(* IEC 61131-3 sources: Lasal-MCP/examples/SampleSource/2_PumpControlSolution/Stations/MachineControl/MachineControl/Class/PumpControl, 1 file *)

(* ---- PumpControl.st ---- *)
(*!
<Class
	Name               = "PumpControl"
	Revision           = "0.0"
	RealtimeTask       = "false"
	CyclicTask         = "true"
	DefCyclictime      = "10 ms"
	BackgroundTask     = "false"
	Sigmatek           = "false"
	OSInterface        = "false"
	HighPriority       = "false"
	Automatic          = "false"
	UpdateMode         = "Prescan"
	SharedCommandTable = "true"
	Objectsize         = "(510,360)">
	<Channels>
		<Server Name="ActFillLevelVisu" Visualized="true" Initialize="false" WriteProtected="true" Retentive="false"/>
		<Server Name="ClassSvr" Visualized="false" Initialize="false" WriteProtected="true" Retentive="false"/>
		<Server Name="MaxBorder" Visualized="true" Initialize="false" WriteProtected="false" Retentive="File"/>
		<Server Name="MinBorder" Visualized="true" Initialize="false" WriteProtected="false" Retentive="File"/>
		<Server Name="PumpVisu" Visualized="true" Initialize="false" WriteProtected="true" Retentive="false"/>
		<Client Name="ActFillLevel" Required="true" Internal="false"/>
		<Client Name="Pump" Required="true" Internal="false"/>
	</Channels>
</Class>
*)
PumpControl : CLASS
  //Servers:
	ClassSvr 	: SvrChCmd_DINT;
	MaxBorder 	: SvrCh_DINT;
	MinBorder 	: SvrCh_DINT;
	PumpVisu 	: SvrCh_DINT;
	ActFillLevelVisu 	: SvrCh_DINT;
  //Clients:
	Pump 	: CltCh_DINT;
	ActFillLevel 	: CltCh_DINT;
  //Variables:
  //Functions:

	FUNCTION VIRTUAL GLOBAL CyWork
		VAR_INPUT
			EAX 	: UDINT;
		END_VAR
		VAR_OUTPUT
			state (EAX) 	: UDINT;
		END_VAR;

	FUNCTION VIRTUAL GLOBAL PumpVisu::Read
		VAR_OUTPUT
			output (EAX) 	: DINT;
		END_VAR;

	FUNCTION VIRTUAL GLOBAL ActFillLevelVisu::Read
		VAR_OUTPUT
			output (EAX) 	: DINT;
		END_VAR;
  //Tables:
	FUNCTION @STD
		VAR_OUTPUT
			ret_code	: CONFSTATES;
		END_VAR;
	FUNCTION GLOBAL TAB @CT_;
END_CLASS;

FUNCTION VIRTUAL GLOBAL PumpControl::CyWork
	VAR_INPUT
		EAX 	: UDINT;
	END_VAR
	VAR_OUTPUT
		state (EAX) 	: UDINT;
	END_VAR

  ActFillLevel := ActFillLevel.Read();

  if ActFillLevel >= MaxBorder then
    Pump := 1;
  elsif ActFillLevel <= MinBorder then
    Pump := 0;
  end_if;

  Pump.Write (Pump);

	state := READY;

END_FUNCTION

FUNCTION VIRTUAL GLOBAL PumpControl::PumpVisu::Read
	VAR_OUTPUT
		output (EAX) 	: DINT;
	END_VAR

	PumpVisu := Pump;

	output := PumpVisu;

END_FUNCTION

FUNCTION VIRTUAL GLOBAL PumpControl::ActFillLevelVisu::Read
	VAR_OUTPUT
		output (EAX) 	: DINT;
	END_VAR

	ActFillLevelVisu := ActFillLevel;

	output := ActFillLevelVisu;

END_FUNCTION
